Fanuc KAREL source: KT00492.KL

PROGRAM KT00492
%NOLOCKGROUP
VAR
  P1: POSITION
  P2: JOINTPOS
  OUT: JOINTPOS
BEGIN
  OUT = P1 : P2
END KT00492
